{attribute 'qualified_only'}
{attribute 'strict'}
TYPE E_UmTutorialState :
(
	NoCmd
);
END_TYPE

(* stored: Version 1.1.0.1, ProductVersion 3.1.4024.12
   DUT E_UmTutorialState: Id {a128ae15-d315-4719-b531-512f438440f7} *)
